# EPICS autosave request: 1.5.0/debian-12/7.0.10/modules/ADCore-ee039d2/db/NDTimeSeries_settings.req
$(P)$(R)TSNumPoints
$(P)$(R)TSTimePerPointLink.DOL
$(P)$(R)TSAveragingTime
$(P)$(R)TSRead.SCAN
$(P)$(R)TSAcquireMode
file "NDPluginBase_settings.req", P=$(P), R=$(R)
